Fanuc KAREL source: KT00395.KL

PROGRAM KT00395
%NOLOCKGROUP
VAR
  P1: JOINTPOS
  P2: POSITION
  OUT: BOOLEAN
BEGIN
  OUT = P1 <= P2
END KT00395
